(* IEC 61131-3 sources: plc-process-lib/tests/GVLs, 7 files *)

(* ---- GVL_TestsAiDi.gvl.st ---- *)
// Назначение: экземпляры наборов тестов семейства входов (FB_AnalogInput, FB_DigitalInput).
//             Объявление экземпляра регистрирует набор в coUnit; PRG_Tests их не перечисляет.
//             {attribute 'linkalways'} обязателен: без него CODESYS 3.5.17 не включает GVL в
//             приложение, и наборы молча не выполняются (docs/TESTING.md).
// Автор:      kr0nsch
// Версия:     0.1.0
// Документ:   docs/TESTING.md
{attribute 'qualified_only'}
{attribute 'linkalways'}
VAR_GLOBAL
    fbAnalogInputTest  : FB_AnalogInput_Test;    // FB_AnalogInput: масштабирование, NE 43, фильтр, уставки, подмена
    fbDigitalInputTest : FB_DigitalInput_Test;   // FB_DigitalInput: задержки, инверсия, подмена, отказ канала
END_VAR

(* ---- GVL_TestsAlarm.gvl.st ---- *)
// Назначение: экземпляры наборов тестов тревог и базы устройств (этап 2 основы) и зондов времени
//             выполнения. Объявление экземпляра регистрирует набор в coUnit; PRG_Tests их не
//             перечисляет. {attribute 'linkalways'} обязателен (docs/TESTING.md).
// Автор:      kr0nsch
// Версия:     0.1.0
// Документ:   docs/TESTING.md
{attribute 'qualified_only'}
{attribute 'linkalways'}
VAR_GLOBAL
    fbAlarmTest      : FB_Alarm_Test;        // FB_Alarm: состояния ISA-18.2, задержки, shelve, подавление, OOS, события
    fbDeviceBaseTest : FB_DeviceBase_Test;   // FB_DeviceBase через FB_TestDevice: режимы, LKG, NE 107, тревоги
    fbRuntimeTest    : FB_Runtime_Test;      // вопросы 24.2 контракта, решаемые тестом на Control Win V3
END_VAR

(* ---- GVL_TestsFoundation.gvl.st ---- *)
// Назначение: экземпляры наборов тестов основы библиотеки (время, утилиты, общие типы).
//             Объявление экземпляра регистрирует набор в coUnit; PRG_Tests их не перечисляет.
//             {attribute 'linkalways'} обязателен: на GVL никто не ссылается, и без атрибута
//             CODESYS 3.5.17 не включает её в приложение — наборы молча не выполняются
//             (проверено зондом, docs/TESTING.md).
// Автор:      kr0nsch
// Версия:     0.1.0
// Документ:   docs/TESTING.md
{attribute 'qualified_only'}
{attribute 'linkalways'}
VAR_GLOBAL
    fbTimeTest   : FB_Time_Test;     // F_LTimeToSec, F_TimeToSec, FB_FakeTime, FB_SystemTime, FB_Delay
    fbUtilTest   : FB_Util_Test;     // F_IsFinite, F_Ne107Worst, F_RateLimit, FB_StartsWindow, FB_LimitMonitor
    fbCommonTest : FB_Common_Test;   // общие типы: SIZEOF, значения по умолчанию, интерфейсы, FB_TestSink
END_VAR

(* ---- GVL_TestsIntegration.gvl.st ---- *)
// Назначение: экземпляр набора межсемейных тестов устройств (все семь типов вместе). Объявление
//             экземпляра регистрирует набор в coUnit; PRG_Tests его не перечисляет.
//             {attribute 'linkalways'} обязателен (docs/TESTING.md).
// Автор:      kr0nsch
// Версия:     0.1.0
// Документ:   docs/TESTING.md, раздел «Межсемейные тесты»
{attribute 'qualified_only'}
{attribute 'linkalways'}
VAR_GLOBAL
    fbIntegrationTest : FB_Integration_Test;   // семь типов устройств: умолчания Cfg, тип, слоты тревог
END_VAR

(* ---- GVL_TestsMotor.gvl.st ---- *)
// Назначение: экземпляры наборов тестов семейства двигателей (FB_Motor, FB_MotorVfd). Объявление
//             экземпляра регистрирует набор в coUnit; PRG_Tests их не перечисляет.
//             {attribute 'linkalways'} обязателен (docs/TESTING.md).
// Автор:      kr0nsch
// Версия:     0.1.0
// Документ:   docs/TESTING.md
{attribute 'qualified_only'}
{attribute 'linkalways'}
VAR_GLOBAL
    fbMotorTest    : FB_Motor_Test;      // FB_Motor: режимы, контроль ОС, отказы, блокировки, времена, счётчики
    fbMotorVfdTest : FB_MotorVfd_Test;   // FB_MotorVfd: задание скорости, связь с ПЧ, рассогласование, интерфейсы
END_VAR

(* ---- GVL_TestsPid.gvl.st ---- *)
// Назначение: экземпляр набора тестов семейства ПИД. Объявление экземпляра регистрирует набор в
//             coUnit; PRG_Tests его не перечисляет. {attribute 'linkalways'} обязателен
//             (docs/TESTING.md).
// Автор:      kr0nsch
// Версия:     0.1.0
// Документ:   docs/fb/FB_PID.md
{attribute 'qualified_only'}
{attribute 'linkalways'}
VAR_GLOBAL
    fbPidTest : FB_Pid_Test;   // FB_PID: алгоритм, anti-windup, режимы, задание, отказ PV, контур с FOPDT
END_VAR

(* ---- GVL_TestsValve.gvl.st ---- *)
// Назначение: экземпляры наборов тестов семейства арматуры (FB_Valve, FB_ControlValve).
//             Объявление экземпляра регистрирует набор в coUnit; PRG_Tests их не перечисляет.
//             {attribute 'linkalways'} обязателен: на GVL никто не ссылается, и без атрибута
//             CODESYS 3.5.17 не включает её в приложение — наборы молча не выполняются
//             (docs/TESTING.md).
// Автор:      kr0nsch
// Версия:     0.1.0
// Документ:   docs/TESTING.md
{attribute 'qualified_only'}
{attribute 'linkalways'}
VAR_GLOBAL
    fbValveTest        : FB_Valve_Test;          // FB_Valve: ход, концевики, реверс, соленоиды, блокировки, режимы
    fbControlValveTest : FB_ControlValve_Test;   // FB_ControlValve: рампа, пределы, рассогласование, безопасность
END_VAR
